// TIA Portal V20 export
// export: Created 2026-10-12T15:52:20.32815Z, ExportSetting WithDefaults, DisplayName Totally Integrated Automation Portal, DisplayVersion V20, DisplayName TIA Portal Openness, DisplayVersion V20, DisplayName TIA Portal Teamcenter Gateway, DisplayVersion V20, DisplayName TIA Portal Version Control Interface, DisplayVersion V20, DisplayName SINAMICS Startdrive Advanced, DisplayVersion V20 SP1 Update 2, DisplayName SINAMICS Startdrive G110M, G120, G120C, G120D, G120P, G115D, DisplayVersion V20 SP1 Update 2, DisplayName SINAMICS Startdrive G130, G150, S120, S150, SINAMICS MV, G220, S200, S210, DisplayVersion V20 SP1 Update 2, DisplayName STEP 7 Professional, DisplayVersion V20, DisplayName STEP 7 Safety, DisplayVersion V20, DisplayName WinCC Basic/Comfort/Advanced, DisplayVersion V20, DisplayName WinCC Professional, DisplayVersion V20, DisplayName WinCC Unified, DisplayVersion V20
FUNCTION "FRK_SetRecord" : Int   // FC114, SCL
{ S7_Optimized_Access := 'TRUE' }
VERSION : 0.1
// stored: AutoNumber true, IsIECCheckEnabled false, SetENOAutomatically false, UDAEnableTagReadback false
   VAR_INPUT
      RootIndex : Int;
      Scope : String;
      WriteKey : String;
   END_VAR
   VAR_TEMP
      Index : Int;
   END_VAR
BEGIN

   #FRK_SetRecord := 0;
   FOR #Index := 1 TO "FRK_SetRuntime".Work[#RootIndex].Payload.Info.RecordCount DO
       IF "FRK_SetRuntime".Work[#RootIndex].Payload.Records[#Index].Scope = #Scope AND "FRK_SetRuntime".Work[#RootIndex].Payload.Records[#Index].WriteKey = #WriteKey THEN
           #FRK_SetRecord := #Index;
           RETURN;
       END_IF;
   END_FOR;
END_FUNCTION
